(* IEC 61131-3 sources: ZPLC/packages/zplc-ide/projects/door_alarm_il_starter/src, 1 file *)

(* ---- DoorAlarm.il ---- *)
PROGRAM DoorAlarm
VAR_INPUT
    Armed AT %I0.0 : BOOL;
    DoorOpen AT %I0.1 : BOOL;
    Silence AT %I0.2 : BOOL;
END_VAR
VAR_OUTPUT
    Siren AT %Q0.0 : BOOL;
END_VAR

        LD    Armed
        AND   DoorOpen
        ST    Siren
END_PROGRAM
